// TIA Portal V21 export
// export: Created 2026-11-21T10:55:36.0525943Z, ExportSetting WithDefaults, DisplayName Totally Integrated Automation Portal, DisplayVersion V21, DisplayName STEP 7 Professional, DisplayVersion V21, DisplayName STEP 7 Safety, DisplayVersion V21, DisplayName Tech WebApplication, DisplayVersion V21, DisplayName WinCC Basic/Comfort/Advanced, DisplayVersion V21, DisplayName WinCC Unified, DisplayVersion V21
VAR_GLOBAL   // PLC tag table "Outputs"
   Infeed_Motor AT %Q0.0 : Bool;   // Infeed conveyor motor
   Outfeed_Motor AT %Q0.1 : Bool;   // Outfeed conveyor motor
   Filler_Valve AT %Q0.2 : Bool;   // Opens the fill valve
   Lamp_Running AT %Q0.3 : Bool;   // The line runs
   Lamp_Fault AT %Q0.4 : Bool;   // A fault waits to be acknowledged
END_VAR
